Yaskawa INFORM job: MAIN_1.JBI

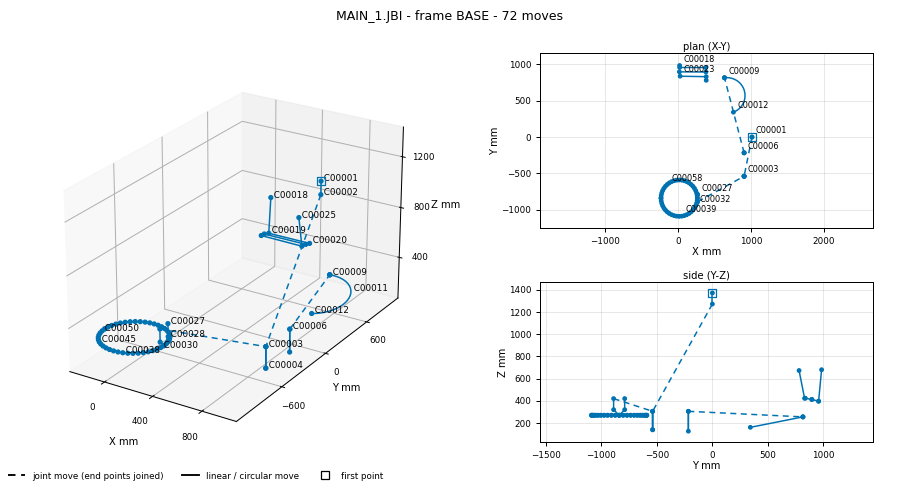
[picture p0: tool path of MAIN_1.JBI in frame BASE, 72 of 80 moves have a stored position in this frame; points joined in program order, loops and branches not executed]
/JOB
//NAME MAIN_1
//POS
///NPOS 80,0,0,0,0,0
///TOOL 9
///POSTYPE PULSE
///PULSE
C00000=0,0,0,0,0,0
///TOOL 9
///POSTYPE BASE
///RECTAN
///RCONF 1,0,0,0,0,0,0,0
C00001=1015.000,0.000,1372.000,0.00,90.00,0.00
///RCONF 0,0,0,0,0,0,0,0
C00002=1015.000,0.000,1272.000,0.00,90.00,0.00
///TOOL 1
///RCONF 1,0,0,0,0,0,0,0
C00003=906.277,-538.516,305.356,-180.00,0.18,180.00
C00004=906.799,-538.504,139.112,180.00,0.18,-180.00
///POSTYPE PULSE
///PULSE
C00005=-29,47,0,27,25,-52
///TOOL 1
///POSTYPE BASE
///RECTAN
///RCONF 1,0,0,0,0,0,0,0
C00006=906.285,-216.481,305.347,-180.00,0.19,180.00
C00007=906.864,-216.486,126.235,-180.00,0.19,180.00
C00008=906.285,-216.481,305.347,-180.00,0.19,180.00
C00009=636.704,815.780,255.156,178.91,11.18,-95.59
C00010=636.704,815.780,255.156,178.91,11.18,-95.59
C00011=884.547,696.689,231.503,178.91,11.18,-95.59
C00012=759.304,342.075,161.073,178.91,11.18,-95.59
///POSTYPE PULSE
///PULSE
C00013=25,41,30,88,29,-142
C00014=39,53,-5,56,30,-93
C00015=52,46,7,67,20,-93
///TOOL 1
///POSTYPE BASE
///RECTAN
///RCONF 1,0,0,0,0,0,0,0
C00016=636.704,815.780,255.156,178.91,11.18,-95.59
///POSTYPE PULSE
///PULSE
C00017=0,0,0,0,0,0
///TOOL 1
///POSTYPE BASE
///RECTAN
///RCONF 1,0,0,0,0,0,0,0
C00018=19.898,984.071,680.331,-179.53,-5.43,-94.93
C00019=19.898,957.021,396.618,-179.53,-5.43,-94.93
C00020=378.402,957.130,396.607,-179.53,-5.43,-94.93
C00021=380.996,895.077,412.492,-178.35,-18.14,-95.29
C00022=16.551,897.073,411.836,-178.35,-18.14,-95.29
C00023=26.434,837.238,423.682,179.59,4.35,-95.46
C00024=385.448,830.764,422.747,178.91,11.18,-95.59
C00025=385.448,781.089,672.861,178.91,11.18,-95.59
///POSTYPE PULSE
///PULSE
C00026=0,0,0,0,0,0
///TOOL 1
///POSTYPE BASE
///RECTAN
///RCONF 1,0,0,0,0,0,0,0
C00027=266.281,-790.141,419.997,-179.97,0.35,-180.00
C00028=266.896,-790.185,319.999,-179.97,0.35,-180.00
C00029=263.637,-840.080,270.000,-179.97,0.35,-180.00
C00030=261.092,-875.659,270.000,-179.93,0.34,-180.00
C00031=253.510,-910.513,270.000,-179.88,0.33,-180.00
C00032=241.045,-943.934,270.000,-179.83,0.31,-180.00
C00033=223.950,-975.240,270.000,-179.79,0.28,-180.00
C00034=202.574,-1003.795,270.000,-179.75,0.25,-180.00
C00035=177.352,-1029.017,270.000,-179.72,0.21,-180.00
C00036=148.797,-1050.393,270.000,-179.69,0.17,-180.00
C00037=117.491,-1067.488,270.000,-179.67,0.12,-180.00
C00038=84.070,-1079.953,270.000,-179.65,0.07,-180.00
C00039=49.216,-1087.535,270.000,-179.65,0.03,-180.00
C00040=13.637,-1090.080,270.000,-179.65,-0.03,-180.00
C00041=-21.942,-1087.535,270.000,-179.65,-0.07,-180.00
C00042=-56.796,-1079.953,270.000,-179.67,-0.12,180.00
C00043=-90.217,-1067.488,270.000,-179.69,-0.17,180.00
C00044=-121.523,-1050.393,270.000,-179.72,-0.21,180.00
C00045=-150.078,-1029.017,270.000,-179.75,-0.25,180.00
C00046=-175.300,-1003.795,270.000,-179.79,-0.28,180.00
C00047=-196.676,-975.240,270.000,-179.83,-0.31,180.00
C00048=-213.771,-943.934,270.000,-179.88,-0.33,180.00
C00049=-226.236,-910.513,270.000,-179.93,-0.35,-180.00
C00050=-233.818,-875.659,270.000,-179.97,-0.35,-180.00
C00051=-236.363,-840.080,270.000,-179.97,-0.35,-180.00
C00052=-236.363,-840.080,270.000,179.97,-0.35,-180.00
C00053=-233.818,-804.501,270.000,179.93,-0.35,-180.00
C00054=-226.236,-769.647,270.000,179.88,-0.33,-180.00
C00055=-213.771,-736.226,270.000,179.83,-0.31,-180.00
C00056=-196.676,-704.920,270.000,179.79,-0.28,-180.00
C00057=-175.300,-676.365,270.000,179.75,-0.25,-180.00
C00058=-150.078,-651.143,270.000,179.72,-0.21,-180.00
C00059=-121.523,-629.767,270.000,179.69,-0.17,-180.00
C00060=-90.217,-612.672,270.000,179.67,-0.12,-180.00
C00061=-56.796,-600.207,270.000,179.65,-0.07,-180.00
C00062=-21.942,-592.625,270.000,179.65,-0.03,-180.00
C00063=13.637,-590.080,270.000,179.65,0.03,-180.00
C00064=49.216,-592.625,270.000,179.66,0.07,-180.00
C00065=84.070,-600.207,270.000,179.67,0.12,180.00
C00066=117.491,-612.672,270.000,179.69,0.17,180.00
C00067=148.797,-629.767,270.000,179.72,0.21,180.00
C00068=177.352,-651.143,270.000,179.75,0.25,180.00
C00069=202.574,-676.365,270.000,179.79,0.28,180.00
C00070=223.950,-704.920,270.000,179.83,0.31,180.00
C00071=241.045,-736.226,270.000,179.88,0.33,180.00
C00072=253.510,-769.647,270.000,179.93,0.35,-180.00
C00073=261.092,-804.501,270.000,179.97,0.35,-180.00
C00074=263.637,-840.080,270.000,179.97,0.35,-180.00
C00075=266.895,-889.975,319.999,179.97,0.35,-180.00
C00076=266.279,-890.019,419.997,179.97,0.35,-180.00
C00077=906.277,-538.516,305.356,-180.00,0.18,180.00
C00078=906.799,-538.504,139.112,180.00,0.18,-180.00
C00079=906.277,-538.516,305.356,-180.00,0.18,180.00
//INST
///DATE 2023/01/01 00:00
///COMM Generated using RoboDK
///ATTR SC,RW,RJ
///GROUP1 RB1
NOP
'Program generated by RoboDK v
'5.6.9 for RoboDK Industrial o
'n 26/02/2024 09:58:20
'Using nominal kinematics.
MOVJ C00000 VJ=50.00
MOVJ C00001 VJ=50.00
MOVL C00002 V=100.0
DOUT OT#(5) ON
DOUT OT#(5) ON
DOUT OT#(5) 0.5
DOUT OT#(5) true
DOUT OT#(5) ON
DOUT OT#(5) ON
DOUT OT#(5) 0.5
DOUT OT#(5) true
DOUT var val
DOUT var val
WAIT IN#(5)=ON
WAIT IN#(5)=ON
WAIT IN#(5)=0.5
WAIT IN#(5)=true
WAIT IN#(5)=ON T=0.10
WAIT var=val
WAIT var=val T=0.10
MSG "Message"
CALL JOB:REMOTE_
CODE_INSERT_172
'Insert Comment
'Using Frame Pick and Place (t
'argets wrt base):
'719.0,-664.0,0.0,0.0,0.0,0.0
'Tool 1 (Tool 1) should be clo
'se to:
'129.1,0.0,85.5,0.0,22.8,0.0
MOVJ C00003 VJ=100.0 ACC=100 DEC=100
MOVL C00004 V=100.0 ACC=100 DEC=100
DOUT OT#(5) ON
CALL JOB:PICK_PA
MOVL C00005 V=300.0 ACC=100 DEC=100
MOVL C00006 V=300.0 ACC=100 DEC=100
'MoveSearch command not implem
'ented
MOVL C00007 V=100.0 ACC=100 DEC=100
DOUT OT#(5) OFF
CALL JOB:PLACE_P
MOVL C00008 V=100.0 ACC=100 DEC=100
'Using Frame Circular (targets
' wrt base):
'577.7,392.2,0.0,0.0,0.0,39.0
MOVJ C00009 VJ=100.0 ACC=100 DEC=100
MOVC C00010 V=100.0 ACC=100 DEC=100 PL=8
MOVC C00011 V=100.0 ACC=100 DEC=100 PL=8
MOVC C00012 V=100.0 ACC=100 DEC=100 PL=8
MOVC C00013 V=100.0 ACC=100 DEC=100 PL=8
MOVC C00014 V=100.0 ACC=100 DEC=100 PL=8
MOVC C00015 V=100.0 ACC=100 DEC=100 PL=8
MOVL C00016 V=100.0 ACC=100 DEC=100
MOVJ C00017 VJ=100.0 ACC=100 DEC=100
'Using Frame Inspection (targe
'ts wrt base):
'0.0,782.7,377.6,0.0,0.0,0.0
MOVJ C00018 VJ=100.0 ACC=100 DEC=100
MOVL C00019 V=100.0 ACC=100 DEC=100
MOVL C00020 V=100.0 ACC=100 DEC=100
MOVL C00021 V=100.0 ACC=100 DEC=100
MOVL C00022 V=100.0 ACC=100 DEC=100
MOVL C00023 V=100.0 ACC=100 DEC=100
MOVL C00024 V=100.0 ACC=100 DEC=100
MOVL C00025 V=100.0 ACC=100 DEC=100
MOVJ C00026 VJ=100.0 ACC=100 DEC=100
CALL JOB:EVENT_P
'Using Frame Inspection (targe
'ts wrt base):
'13.6,-840.1,0.0,0.0,0.0,-90.0
'Show Tool 1
MOVJ C00027 VJ=100.0 ACC=100 DEC=100
CALL JOB:EVENT_P
MOVL C00028 V=1000.0 ACC=100 DEC=100
MOVL C00029 V=1000.0 ACC=100 DEC=100
CALL JOB:EVENT_P
MOVL C00030 V=50.0 ACC=100 DEC=100
MOVL C00031 V=50.0 ACC=100 DEC=100
MOVL C00032 V=50.0 ACC=100 DEC=100
MOVL C00033 V=50.0 ACC=100 DEC=100
MOVL C00034 V=50.0 ACC=100 DEC=100
MOVL C00035 V=50.0 ACC=100 DEC=100
MOVL C00036 V=50.0 ACC=100 DEC=100
MOVL C00037 V=50.0 ACC=100 DEC=100
MOVL C00038 V=50.0 ACC=100 DEC=100
MOVL C00039 V=50.0 ACC=100 DEC=100
MOVL C00040 V=50.0 ACC=100 DEC=100
MOVL C00041 V=50.0 ACC=100 DEC=100
MOVL C00042 V=50.0 ACC=100 DEC=100
MOVL C00043 V=50.0 ACC=100 DEC=100
MOVL C00044 V=50.0 ACC=100 DEC=100
MOVL C00045 V=50.0 ACC=100 DEC=100
MOVL C00046 V=50.0 ACC=100 DEC=100
MOVL C00047 V=50.0 ACC=100 DEC=100
MOVL C00048 V=50.0 ACC=100 DEC=100
MOVL C00049 V=50.0 ACC=100 DEC=100
MOVL C00050 V=50.0 ACC=100 DEC=100
MOVL C00051 V=50.0 ACC=100 DEC=100
MOVL C00052 V=50.0 ACC=100 DEC=100
MOVL C00053 V=50.0 ACC=100 DEC=100
MOVL C00054 V=50.0 ACC=100 DEC=100
MOVL C00055 V=50.0 ACC=100 DEC=100
MOVL C00056 V=50.0 ACC=100 DEC=100
MOVL C00057 V=50.0 ACC=100 DEC=100
MOVL C00058 V=50.0 ACC=100 DEC=100
MOVL C00059 V=50.0 ACC=100 DEC=100
MOVL C00060 V=50.0 ACC=100 DEC=100
MOVL C00061 V=50.0 ACC=100 DEC=100
MOVL C00062 V=50.0 ACC=100 DEC=100
MOVL C00063 V=50.0 ACC=100 DEC=100
MOVL C00064 V=50.0 ACC=100 DEC=100
MOVL C00065 V=50.0 ACC=100 DEC=100
MOVL C00066 V=50.0 ACC=100 DEC=100
MOVL C00067 V=50.0 ACC=100 DEC=100
MOVL C00068 V=50.0 ACC=100 DEC=100
MOVL C00069 V=50.0 ACC=100 DEC=100
MOVL C00070 V=50.0 ACC=100 DEC=100
MOVL C00071 V=50.0 ACC=100 DEC=100
MOVL C00072 V=50.0 ACC=100 DEC=100
MOVL C00073 V=50.0 ACC=100 DEC=100
MOVL C00074 V=50.0 ACC=100 DEC=100
CALL JOB:EVENT_P
MOVL C00075 V=1000.0 ACC=100 DEC=100
MOVL C00076 V=1000.0 ACC=100 DEC=100
CALL JOB:EVENT_P
CALL JOB:EVENT_P
'Using Frame Pick and Place (t
'argets wrt base):
'719.0,-664.0,0.0,0.0,0.0,0.0
MOVJ C00077 VJ=100.0 ACC=100 DEC=100
TIMER T=1.25
MOVL C00078 V=1000.0 ACC=100 DEC=100
WAIT IN#(1)=ON
MOVL C00079 V=1000.0 ACC=100 DEC=100
CALL JOB:PROG1_W
END
